        string sFontStyle
        string sFontWeight
        string sTextAlignment
public utLabel utLbl_Axis_Data
  [0]
    utAppearance Appearance
      [0]
        bool bVisibility
        string sBackgroundColour = "#FFFFFF"
        string sColour
    utBorder Border
      [0]
        num nBorderWidth
        string sBorderColour
        string sBorderStyle
    utCommon Common
      [0]
        string sID = "lbl_Axis_Data"
        string sPage = "Disk://SmartTCP_CS9/tx2/interface/Page_Main"
        string sText = "6轴"
    utData Data
      [0]
        bool bStatus
        num nVal = 99
    utEvents Events
      [0]
        bool bClick
        bool bMouseDown
        bool bMouseUp
    utText Text
      [0]
        num nFontSize
        string sFontFamily
        string sFontStyle
        string sFontWeight
        string sTextAlignment
public utLabel utLbl_CheckBox_a[3]
  [0]
    utAppearance Appearance
      [0]
        bool bVisibility
        string sBackgroundColour = "#FFFFFF"
        string sColour
    utBorder Border
      [0]
        num nBorderWidth
        string sBorderColour
        string sBorderStyle
    utCommon Common
      [0]
        string sID = "lbl_CheckBox_a0"
        string sPage = "Disk://SmartTCP_CS9/tx2/interface/Page_Container_Main"
        string sText = "3点标定"
    utData Data
      [0]
        bool bStatus
        num nVal = 99
    utEvents Events
      [0]
        bool bClick
        bool bMouseDown
        bool bMouseUp
    utText Text
      [0]
        num nFontSize
        string sFontFamily
        string sFontStyle
        string sFontWeight
        string sTextAlignment
  [1]
    utAppearance Appearance
      [0]
        bool bVisibility
        string sBackgroundColour = "#FFFFFF"
        string sColour
    utBorder Border
      [0]
        num nBorderWidth
        string sBorderColour
        string sBorderStyle
    utCommon Common
      [0]
        string sID = "lbl_CheckBox_a1"
        string sPage = "Disk://SmartTCP_CS9/tx2/interface/Page_Container_Main"
        string sText = "4点标定"
    utData Data
      [0]
        bool bStatus
        num nVal = 99
    utEvents Events
      [0]
        bool bClick = true
        bool bMouseDown
        bool bMouseUp
    utText Text
      [0]
        num nFontSize
        string sFontFamily
        string sFontStyle
        string sFontWeight
        string sTextAlignment
  [2]
    utAppearance Appearance
      [0]
        bool bVisibility
        string sBackgroundColour = "#FFFFFF"
        string sColour
    utBorder Border
      [0]
        num nBorderWidth
        string sBorderColour
        string sBorderStyle
    utCommon Common
      [0]
        string sID = "lbl_CheckBox_a2"
        string sPage = "Disk://SmartTCP_CS9/tx2/interface/Page_Container_Main"
        string sText = "7点标定"
    utData Data
      [0]
        bool bStatus
        num nVal = 99
    utEvents Events
      [0]
        bool bClick
        bool bMouseDown
        bool bMouseUp
    utText Text
      [0]
        num nFontSize
        string sFontFamily
        string sFontStyle
        string sFontWeight
        string sTextAlignment
public utLabel utLbl_CheckBox_b[2]
  [0]
    utAppearance Appearance
      [0]
        bool bVisibility
        string sBackgroundColour = "#FFFFFF"
        string sColour
    utBorder Border
      [0]
        num nBorderWidth
        string sBorderColour
        string sBorderStyle
    utCommon Common
      [0]
        string sID = "lbl_CheckBox_b0"
        string sPage = "Disk://SmartTCP_CS9/tx2/interface/Page_Container_Main"
        string sText = "2点180°"
    utData Data
      [0]
        bool bStatus
        num nVal = 99
    utEvents Events
      [0]
        bool bClick
        bool bMouseDown
        bool bMouseUp
    utText Text
      [0]
        num nFontSize
        string sFontFamily
        string sFontStyle
        string sFontWeight
        string sTextAlignment
  [1]
    utAppearance Appearance
      [0]
        bool bVisibility
        string sBackgroundColour = "#FFFFFF"
        string sColour
    utBorder Border
      [0]
        num nBorderWidth
        string sBorderColour
        string sBorderStyle
    utCommon Common
      [0]
        string sID = "lbl_CheckBox_b1"
        string sPage = "Disk://SmartTCP_CS9/tx2/interface/Page_Container_Main"
        string sText = "3点120°"
    utData Data
      [0]
        bool bStatus
        num nVal = 99
    utEvents Events
      [0]
        bool bClick
        bool bMouseDown
        bool bMouseUp
    utText Text
      [0]
        num nFontSize
        string sFontFamily
        string sFontStyle
        string sFontWeight
        string sTextAlignment
public utLabel utLbl_CurrentPos_Data[6]
  [0]
    utAppearance Appearance
      [0]
        bool bVisibility
        string sBackgroundColour = "#FFFFFF"
        string sColour
    utBorder Border
      [0]
        num nBorderWidth
        string sBorderColour
        string sBorderStyle
    utCommon Common
      [0]
        string sID = "lbl_CurrentPos_Data0"
        string sPage = "Disk://SmartTCP_CS9/tx2/interface/Page_Main"
        string sText = "1137.12 "
    utData Data
      [0]
        bool bStatus
        num nVal = 99
    utEvents Events
      [0]
        bool bClick
        bool bMouseDown
        bool bMouseUp
    utText Text
      [0]
        num nFontSize
        string sFontFamily
        string sFontStyle
        string sFontWeight
        string sTextAlignment
  [1]
    utAppearance Appearance
      [0]
        bool bVisibility
        string sBackgroundColour = "#FFFFFF"
        string sColour
    utBorder Border
      [0]
        num nBorderWidth
        string sBorderColour
        string sBorderStyle
    utCommon Common
      [0]
        string sID = "lbl_CurrentPos_Data1"
        string sPage = "Disk://SmartTCP_CS9/tx2/interface/Page_Main"
        string sText = "-108.577"
    utData Data
      [0]
        bool bStatus
        num nVal = 99
    utEvents Events
      [0]
        bool bClick
        bool bMouseDown
        bool bMouseUp
    utText Text
      [0]
        num nFontSize
        string sFontFamily
        string sFontStyle
        string sFontWeight
        string sTextAlignment
  [2]
    utAppearance Appearance
      [0]
        bool bVisibility
        string sBackgroundColour = "#FFFFFF"
        string sColour
    utBorder Border
      [0]
        num nBorderWidth
        string sBorderColour
        string sBorderStyle
    utCommon Common
      [0]
        string sID = "lbl_CurrentPos_Data2"
        string sPage = "Disk://SmartTCP_CS9/tx2/interface/Page_Main"
        string sText = "-202.363"
    utData Data
      [0]
        bool bStatus
        num nVal = 99
    utEvents Events
      [0]
        bool bClick
        bool bMouseDown
        bool bMouseUp
    utText Text
      [0]
        num nFontSize
        string sFontFamily
        string sFontStyle
        string sFontWeight
        string sTextAlignment
  [3]
    utAppearance Appearance
      [0]
        bool bVisibility
        string sBackgroundColour = "#FFFFFF"
        string sColour
    utBorder Border
      [0]
        num nBorderWidth
        string sBorderColour
        string sBorderStyle
    utCommon Common
      [0]
        string sID = "lbl_CurrentPos_Data3"
        string sPage = "Disk://SmartTCP_CS9/tx2/interface/Page_Main"
        string sText = "-0    "
    utData Data
      [0]
        bool bStatus
        num nVal = 99
    utEvents Events
      [0]
        bool bClick
        bool bMouseDown
        bool bMouseUp
    utText Text
      [0]
        num nFontSize
        string sFontFamily
        string sFontStyle
        string sFontWeight
        string sTextAlignment
  [4]
    utAppearance Appearance
      [0]
        bool bVisibility
        string sBackgroundColour = "#FFFFFF"
        string sColour
    utBorder Border
      [0]
        num nBorderWidth
        string sBorderColour
        string sBorderStyle
    utCommon Common
      [0]
        string sID = "lbl_CurrentPos_Data4"
        string sPage = "Disk://SmartTCP_CS9/tx2/interface/Page_Main"
        string sText = "0    "
    utData Data
      [0]
        bool bStatus
        num nVal = 99
    utEvents Events
      [0]
        bool bClick
        bool bMouseDown
        bool bMouseUp
    utText Text
      [0]
        num nFontSize
        string sFontFamily
        string sFontStyle
        string sFontWeight
        string sTextAlignment
  [5]
    utAppearance Appearance
      [0]
        bool bVisibility
        string sBackgroundColour = "#FFFFFF"
        string sColour
    utBorder Border
      [0]
        num nBorderWidth
        string sBorderColour
        string sBorderStyle
    utCommon Common
      [0]
        string sID = "lbl_CurrentPos_Data5"
        string sPage = "Disk://SmartTCP_CS9/tx2/interface/Page_Main"
        string sText = "0.785"
    utData Data
      [0]
        bool bStatus
        num nVal = 99
    utEvents Events
      [0]
        bool bClick
        bool bMouseDown
        bool bMouseUp
    utText Text
      [0]
        num nFontSize
        string sFontFamily
        string sFontStyle
        string sFontWeight
        string sTextAlignment
public utLabel utLbl_CurrentPos_Name[6]
  [0]
    utAppearance Appearance
      [0]
        bool bVisibility
        string sBackgroundColour = "#FFFFFF"
        string sColour
    utBorder Border
      [0]
        num nBorderWidth
        string sBorderColour
        string sBorderStyle
    utCommon Common
      [0]
        string sID = "lbl_CurrentPos_Name0"
        string sPage = "Disk://SmartTCP_CS9/tx2/interface/Page_Main"
        string sText = "X:"
    utData Data
      [0]
        bool bStatus
        num nVal = 99
    utEvents Events
      [0]
        bool bClick
        bool bMouseDown
        bool bMouseUp
    utText Text
      [0]
        num nFontSize
        string sFontFamily
        string sFontStyle
        string sFontWeight
        string sTextAlignment
  [1]
    utAppearance Appearance
      [0]
        bool bVisibility
        string sBackgroundColour = "#FFFFFF"
        string sColour
    utBorder Border
      [0]
        num nBorderWidth
        string sBorderColour
        string sBorderStyle
    utCommon Common
      [0]
        string sID = "lbl_CurrentPos_Name1"
        string sPage = "Disk://SmartTCP_CS9/tx2/interface/Page_Main"
        string sText = "Y:"
    utData Data
      [0]
        bool bStatus
        num nVal = 99
    utEvents Events
      [0]
        bool bClick
        bool bMouseDown
        bool bMouseUp
    utText Text
      [0]
        num nFontSize
        string sFontFamily
        string sFontStyle
        string sFontWeight
        string sTextAlignment
  [2]
    utAppearance Appearance
      [0]
        bool bVisibility
        string sBackgroundColour = "#FFFFFF"
        string sColour
    utBorder Border
      [0]
        num nBorderWidth
        string sBorderColour
        string sBorderStyle
    utCommon Common
      [0]
        string sID = "lbl_CurrentPos_Name2"
        string sPage = "Disk://SmartTCP_CS9/tx2/interface/Page_Main"
        string sText = "Z:"
    utData Data
      [0]
        bool bStatus
        num nVal = 99
    utEvents Events
      [0]
        bool bClick
        bool bMouseDown
        bool bMouseUp
    utText Text
      [0]
        num nFontSize
        string sFontFamily
        string sFontStyle
        string sFontWeight
        string sTextAlignment
  [3]
    utAppearance Appearance
      [0]
        bool bVisibility
        string sBackgroundColour = "#FFFFFF"
        string sColour
    utBorder Border
      [0]
        num nBorderWidth
        string sBorderColour
        string sBorderStyle
    utCommon Common
      [0]
        string sID = "lbl_CurrentPos_Name3"
        string sPage = "Disk://SmartTCP_CS9/tx2/interface/Page_Main"
        string sText = "RX:"
    utData Data
      [0]
        bool bStatus
        num nVal = 99
    utEvents Events
      [0]
        bool bClick
        bool bMouseDown
        bool bMouseUp
    utText Text
      [0]
        num nFontSize
        string sFontFamily
        string sFontStyle
        string sFontWeight
        string sTextAlignment
  [4]
    utAppearance Appearance
      [0]
        bool bVisibility
        string sBackgroundColour = "#FFFFFF"
        string sColour
    utBorder Border
      [0]
        num nBorderWidth
        string sBorderColour
        string sBorderStyle
    utCommon Common
      [0]
        string sID = "lbl_CurrentPos_Name4"
        string sPage = "Disk://SmartTCP_CS9/tx2/interface/Page_Main"
        string sText = "RY:"
    utData Data
      [0]
        bool bStatus
        num nVal = 99
    utEvents Events
      [0]
        bool bClick
        bool bMouseDown
        bool bMouseUp
    utText Text
      [0]
        num nFontSize
        string sFontFamily
        string sFontStyle
        string sFontWeight
        string sTextAlignment
  [5]
    utAppearance Appearance
      [0]
        bool bVisibility
        string sBackgroundColour = "#FFFFFF"
        string sColour
    utBorder Border
      [0]
        num nBorderWidth
        string sBorderColour
        string sBorderStyle
    utCommon Common
      [0]
        string sID = "lbl_CurrentPos_Name5"
        string sPage = "Disk://SmartTCP_CS9/tx2/interface/Page_Main"
        string sText = "RZ:"
    utData Data
      [0]
        bool bStatus
        num nVal = 99
    utEvents Events
      [0]
        bool bClick
        bool bMouseDown
        bool bMouseUp
    utText Text
      [0]
        num nFontSize
        string sFontFamily
        string sFontStyle
        string sFontWeight
        string sTextAlignment
public utLabel utLbl_Info0
  [0]
    utAppearance Appearance
      [0]
        bool bVisibility
        string sBackgroundColour = "#FFFFFF"
        string sColour
    utBorder Border
      [0]
        num nBorderWidth
        string sBorderColour
        string sBorderStyle
    utCommon Common
      [0]
        string sID = "lbl_info0"
        string sPage = "Disk://SmartTCP_CS9/tx2/interface/Page_Main"
        string sText = "操作提醒："
    utData Data
      [0]
        bool bStatus
        num nVal = 101
    utEvents Events
      [0]
        bool bClick
        bool bMouseDown
        bool bMouseUp
    utText Text
      [0]
        num nFontSize
        string sFontFamily
        string sFontStyle
        string sFontWeight
        string sTextAlignment
public utLabel utLbl_Info1
  [0]
    utAppearance Appearance
      [0]
        bool bVisibility
        string sBackgroundColour = "#FFFFFF"
        string sColour
    utBorder Border
      [0]
        num nBorderWidth
        string sBorderColour
        string sBorderStyle
    utCommon Common
      [0]
        string sID = "lbl_info1"
        string sPage = "Disk://SmartTCP_CS9/tx2/interface/Page_Main"
        string sText = "1.旋转TCP(RZ)接近一侧极限"
    utData Data
      [0]
        bool bStatus
        num nVal = 113
    utEvents Events
      [0]
        bool bClick
        bool bMouseDown
        bool bMouseUp
    utText Text
      [0]
        num nFontSize
        string sFontFamily
        string sFontStyle
        string sFontWeight
        string sTextAlignment
public utLabel utLbl_Info2
  [0]
    utAppearance Appearance
      [0]
        bool bVisibility
        string sBackgroundColour = "#FFFFFF"
        string sColour
    utBorder Border
      [0]
        num nBorderWidth
        string sBorderColour
        string sBorderStyle
    utCommon Common
      [0]
        string sID = "lbl_info2"
        string sPage = "Disk://SmartTCP_CS9/tx2/interface/Page_Main"
        string sText = "2.工具垂直姿态对准尖点并记录"
    utData Data
      [0]
        bool bStatus
        num nVal = 102
    utEvents Events
      [0]
        bool bClick = true
        bool bMouseDown
        bool bMouseUp
    utText Text
      [0]
        num nFontSize
        string sFontFamily
        string sFontStyle
        string sFontWeight
        string sTextAlignment
public utLabel utLbl_Info3
  [0]
    utAppearance Appearance
      [0]
        bool bVisibility
        string sBackgroundColour = "#FFFFFF"
        string sColour
    utBorder Border
      [0]
        num nBorderWidth
        string sBorderColour
        string sBorderStyle
    utCommon Common
      [0]
        string sID = "lbl_info3"
        string sPage = "Disk://SmartTCP_CS9/tx2/interface/Page_Main"
        string sText = "3.确保TCP(RZ) 可以反向旋转180°"
    utData Data
      [0]
        bool bStatus
        num nVal = 111
    utEvents Events
      [0]
        bool bClick
        bool bMouseDown
        bool bMouseUp
    utText Text
      [0]
        num nFontSize
        string sFontFamily
        string sFontStyle
        string sFontWeight
        string sTextAlignment
public utLabel utLbl_Info4
  [0]
    utAppearance Appearance
      [0]
        bool bVisibility
        string sBackgroundColour = "#FFFFFF"
        string sColour
    utBorder Border
      [0]
        num nBorderWidth
        string sBorderColour
        string sBorderStyle
    utCommon Common
      [0]
        string sID = "lbl_info4"
        string sPage = "Disk://SmartTCP_CS9/tx2/interface/Page_Main"
        string sText = "4.按记录按钮保存当前位置"
    utData Data
      [0]
        bool bStatus
        num nVal = 105
    utEvents Events
      [0]
        bool bClick = true
        bool bMouseDown
        bool bMouseUp
    utText Text
      [0]
        num nFontSize
        string sFontFamily
        string sFontStyle
        string sFontWeight
        string sTextAlignment
public utLabel utLbl_Language
  [0]
    utAppearance Appearance
      [0]
        bool bVisibility
        string sBackgroundColour = "#FFFFFF"
        string sColour
    utBorder Border
      [0]
        num nBorderWidth
        string sBorderColour
        string sBorderStyle
    utCommon Common
      [0]
        string sID = "lbl_Language"
        string sPage = "Disk://SmartTCP_CS9/tx2/interface/Page_Main"
        string sText = "语言："
    utData Data
      [0]
        bool bStatus
        num nVal = 99
    utEvents Events
      [0]
        bool bClick = true
        bool bMouseDown
        bool bMouseUp
    utText Text
      [0]
        num nFontSize
        string sFontFamily
        string sFontStyle
        string sFontWeight
        string sTextAlignment
public utLabel utLbl_Mounting
  [0]
    utAppearance Appearance
      [0]
        bool bVisibility
        string sBackgroundColour = "#FFFFFF"
        string sColour
    utBorder Border
      [0]
        num nBorderWidth
        string sBorderColour
        string sBorderStyle
    utCommon Common
      [0]
        string sID = "lbl_Mounting"
        string sPage = "Disk://SmartTCP_CS9/tx2/interface/Page_Main"
        string sText = "安装："
    utData Data
      [0]
        bool bStatus
        num nVal = 99
    utEvents Events
      [0]
        bool bClick
        bool bMouseDown
        bool bMouseUp
    utText Text
      [0]
        num nFontSize
        string sFontFamily
        string sFontStyle
        string sFontWeight
        string sTextAlignment
public utLabel utLbl_Offset
  [0]
    utAppearance Appearance
      [0]
        bool bVisibility
        string sBackgroundColour = "#FFFFFF"
        string sColour
    utBorder Border
      [0]
        num nBorderWidth
        string sBorderColour
        string sBorderStyle
    utCommon Common
      [0]
        string sID = "lbl_Offset"
        string sPage = "Disk://SmartTCP_CS9/tx2/interface/Page_Container_Test"
        string sText = "工具补偿："
    utData Data
      [0]
        bool bStatus
        num nVal = 99
    utEvents Events
      [0]
        bool bClick
        bool bMouseDown
        bool bMouseUp
    utText Text
      [0]
        num nFontSize
        string sFontFamily
        string sFontStyle
        string sFontWeight
        string sTextAlignment
public utLabel utLbl_Point
  [0]
    utAppearance Appearance
      [0]
        bool bVisibility
        string sBackgroundColour = "#7CFA3F"
        string sColour
    utBorder Border
      [0]
        num nBorderWidth
        string sBorderColour
        string sBorderStyle
    utCommon Common
      [0]
        string sID = "lbl_Point"
        string sPage = "Disk://SmartTCP_CS9/tx2/interface/Page_Container_Teach"
        string sText = "点位：P1"
    utData Data
      [0]
        bool bStatus
        num nVal = 99
    utEvents Events
      [0]
        bool bClick
        bool bMouseDown
        bool bMouseUp
    utText Text
      [0]
        num nFontSize
        string sFontFamily
        string sFontStyle
        string sFontWeight
        string sTextAlignment
public utLabel utLbl_PosValue_Data[6]
  [0]
    utAppearance Appearance
      [0]
        bool bVisibility
        string sBackgroundColour = "#FFFFFF"
        string sColour
    utBorder Border
      [0]
        num nBorderWidth
        string sBorderColour
        string sBorderStyle
    utCommon Common
      [0]
        string sID = "utLbl_PosValue_Data0"
        string sPage = "Disk://SmartTCP_CS9/tx2/interface/Page_Container_Teach"
        string sText = "1137.12 "
    utData Data
      [0]
        bool bStatus
        num nVal = 99
    utEvents Events
      [0]
        bool bClick
        bool bMouseDown
        bool bMouseUp
    utText Text
      [0]
        num nFontSize
        string sFontFamily
        string sFontStyle
        string sFontWeight
        string sTextAlignment
  [1]
    utAppearance Appearance
      [0]
        bool bVisibility
        string sBackgroundColour = "#FFFFFF"
        string sColour
    utBorder Border
      [0]
        num nBorderWidth
        string sBorderColour
        string sBorderStyle
    utCommon Common
      [0]
        string sID = "utLbl_PosValue_Data1"
        string sPage = "Disk://SmartTCP_CS9/tx2/interface/Page_Container_Teach"
        string sText = "-108.577"
    utData Data
      [0]
        bool bStatus
        num nVal = 99
    utEvents Events
      [0]
        bool bClick
        bool bMouseDown
        bool bMouseUp
    utText Text
      [0]
        num nFontSize
        string sFontFamily
        string sFontStyle
        string sFontWeight
        string sTextAlignment
  [2]
    utAppearance Appearance
      [0]
        bool bVisibility
        string sBackgroundColour = "#FFFFFF"
        string sColour
    utBorder Border
      [0]
        num nBorderWidth
        string sBorderColour
        string sBorderStyle
    utCommon Common
      [0]
        string sID = "utLbl_PosValue_Data2"
        string sPage = "Disk://SmartTCP_CS9/tx2/interface/Page_Container_Teach"
        string sText = "-202.363"
    utData Data
      [0]
        bool bStatus
        num nVal = 99
    utEvents Events
      [0]
        bool bClick
        bool bMouseDown
        bool bMouseUp
    utText Text
      [0]
        num nFontSize
        string sFontFamily
        string sFontStyle
        string sFontWeight
        string sTextAlignment
  [3]
    utAppearance Appearance
      [0]
        bool bVisibility
        string sBackgroundColour = "#FFFFFF"
        string sColour
    utBorder Border
      [0]
        num nBorderWidth
        string sBorderColour
        string sBorderStyle
    utCommon Common
      [0]
        string sID = "utLbl_PosValue_Data3"
        string sPage = "Disk://SmartTCP_CS9/tx2/interface/Page_Container_Teach"
        string sText = "-0    "
    utData Data
      [0]
        bool bStatus
        num nVal = 99
    utEvents Events
      [0]
        bool bClick
        bool bMouseDown
        bool bMouseUp
    utText Text
      [0]
        num nFontSize
        string sFontFamily
        string sFontStyle
        string sFontWeight
        string sTextAlignment
  [4]
    utAppearance Appearance
      [0]
        bool bVisibility
        string sBackgroundColour = "#FFFFFF"
        string sColour
    utBorder Border
      [0]
        num nBorderWidth
        string sBorderColour
        string sBorderStyle
    utCommon Common
      [0]
        string sID = "utLbl_PosValue_Data4"
        string sPage = "Disk://SmartTCP_CS9/tx2/interface/Page_Container_Teach"
        string sText = "0    "
    utData Data
      [0]
        bool bStatus
        num nVal = 99
    utEvents Events
      [0]
        bool bClick
        bool bMouseDown
        bool bMouseUp
    utText Text
      [0]
        num nFontSize
        string sFontFamily
        string sFontStyle
        string sFontWeight
        string sTextAlignment
  [5]
    utAppearance Appearance
      [0]
        bool bVisibility
        string sBackgroundColour = "#FFFFFF"
        string sColour
    utBorder Border
      [0]
        num nBorderWidth
        string sBorderColour
        string sBorderStyle
    utCommon Common
      [0]
        string sID = "utLbl_PosValue_Data5"
        string sPage = "Disk://SmartTCP_CS9/tx2/interface/Page_Container_Teach"
        string sText = "0.785"
    utData Data
      [0]
        bool bStatus
        num nVal = 99
    utEvents Events
      [0]
        bool bClick
        bool bMouseDown
        bool bMouseUp
    utText Text
      [0]
        num nFontSize
        string sFontFamily
        string sFontStyle
        string sFontWeight
        string sTextAlignment
public utLabel utLbl_Step
  [0]
    utAppearance Appearance
      [0]
        bool bVisibility
        string sBackgroundColour = "#FFFFFF"
        string sColour
    utBorder Border
      [0]
        num nBorderWidth
        string sBorderColour
        string sBorderStyle
    utCommon Common
      [0]
        string sID = "lbl_Step"
        string sPage = "Disk://SmartTCP_CS9/tx2/interface/Page_Container_Teach"
        string sText = "步骤：1/2"
    utData Data
      [0]
        bool bStatus
        num nVal = 99
    utEvents Events
      [0]
        bool bClick = true
        bool bMouseDown
        bool bMouseUp
    utText Text
      [0]
        num nFontSize
        string sFontFamily
        string sFontStyle
        string sFontWeight
        string sTextAlignment
public utLabel utLbl_SubTitle1
  [0]
    utAppearance Appearance
      [0]
        bool bVisibility
        string sBackgroundColour = "#FFFFFF"
        string sColour
    utBorder Border
      [0]
        num nBorderWidth
        string sBorderColour
        string sBorderStyle
    utCommon Common
      [0]
        string sID = "lbl_SubTitle1"
        string sPage
        string sText = "版本: V1.0 "
    utData Data
      [0]
        bool bStatus
        num nVal = 5
    utEvents Events
      [0]
        bool bClick
        bool bMouseDown
        bool bMouseUp
    utText Text
      [0]
        num nFontSize
        string sFontFamily
        string sFontStyle
        string sFontWeight
        string sTextAlignment
public utLabel utLbl_SubTitle2
  [0]
    utAppearance Appearance
      [0]
        bool bVisibility
        string sBackgroundColour = "#FFFFFF"
        string sColour
    utBorder Border
      [0]
        num nBorderWidth
        string sBorderColour
        string sBorderStyle
    utCommon Common
      [0]
        string sID = "lbl_SubTitle2"
        string sPage
        string sText = "日期: 2019.11.06"
    utData Data
      [0]
        bool bStatus
        num nVal = 6
    utEvents Events
      [0]
        bool bClick
